TEXTLIST TextList_Piston_Recipe_State
  0 = ' '
  1 = 'Open'
  2 = 'Close'
   = ''
END_TEXTLIST

(* stored: Version 1.1.0.1, ProductVersion 3.1.4024.12
   TextList TextList_Piston_Recipe_State: Id {9f9ac3ce-bd49-47d3-a364-677c4ebcfe58} *)
